Fanuc KAREL source: kc00032.KL

-- PROVISIONAL review KL for V1013-1; original PC SHA256 b398271479e37a14915c29aabffb81e357830e60123dc13346092431d872d32f
-- Incomplete behavior may be omitted. Consult companion uncertainty JSON. Do not deploy.
PROGRAM KC00032
%NOLOCKGROUP
BEGIN
  -- UNRESOLVED_PC offsets 5-55; opcodes 27,22,2A,22,22,22,22,22,22,27,9D,31
  -- UNRESOLVED_PC offsets 60-64; opcodes 7F
END KC00032
